// TIA Portal V21 export
TextList "TL_Bay"  ListRange=Decimal
  TextListEntry   Text="0 BROD"
  TextListEntry   From=1, To=1, Text="1 SKLADIŠTE"
